PROGRAM PRG_TEST
VAR
    fbBendKinematics_Test : FB_BendKinematics_Test;
END_VAR

TcUnit.RUN();

END_PROGRAM

(* stored: Version 1.1.0.1
   POU PRG_TEST: Id {01b11869-cb05-4f63-8eac-354a5879d56a}, SpecialFunc None *)
